(* PLC project PR_TabTrimSeq_Soft2.0 1_workflow_23a3c5_PLC, SiemensToBackhoff Siemens TIA Portal → Beckhoff TwinCAT PLCopen Converter 2.2 *)
(* stored: creationDateTime 2026-10-12T09:25:37.624382, modificationDateTime 2026-10-12T09:25:37.624382 *)

FUNCTION_BLOCK PR_TabTrimSeq_Soft2.0 1_workflow_23a3c5
VAR_INPUT
	iAbort : BOOL;
	iAutoRunning : BOOL;
	iFaultReset : BOOL;
	iPartNotWorkable : BOOL;
	iPartWorkable : BOOL;
	iRFReadDone : BOOL;
	iRFReadError : BOOL;
	iRFWriteDone : BOOL;
	iRFWriteError : BOOL;
	iReject : BOOL;
	iReset_fault : BOOL;
	iRetry : BOOL;
	iRetryCount : INT;
	iSstMode : BOOL;
	iSstPB : BOOL;
	iStartFrmFibro : BOOL;
	iStartFrmFibroSeq : BOOL;
	iTrimOver : BOOL;
	iZAxisDownOver : BOOL;
	iZAxisUpOver : BOOL;
END_VAR
VAR_OUTPUT
	qError : ARRAY[0..2] OF BOOL;
	qMessage : ARRAY[0..2] OF BOOL;
	qScrapSuction : BOOL;
	qTrimOprnOver : BOOL;
	qTrimStartCmd : BOOL;
	qZAxisUp : BOOL;
	qzAxisDown : BOOL;
END_VAR
VAR
	c20_ChkRecovery_T1 : BOOL;
	c20_ChkRecovery_T2 : BOOL;
	c20_ChkRecovery_T3 : BOOL;
	c21_WtRFIDReadOver_T1 : BOOL;
	c21_WtRFIDReadOver_T2 : BOOL;
	c22_ChkRetryCountRead_T1 : BOOL;
	c22_ChkRetryCountRead_T2 : BOOL;
	c23_WtOpDecisionRead_T1 : BOOL;
	c23_WtOpDecisionRead_T2 : BOOL;
	c24_ChkPartWorkable_T1 : BOOL;
	c24_ChkPartWorkable_T2 : BOOL;
	c61_WtRFIDWriteOver_T1 : BOOL;
	c61_WtRFIDWriteOver_T2 : BOOL;
	c62_ChkRetryCountWrite_T1 : BOOL;
	c62_ChkRetryCountWrite_T2 : BOOL;
	c63_WtOpDecisionWrite_T1 : BOOL;
	c63_WtOpDecisionWrite_T2 : BOOL;
	StateNo : INT;
	s10_WtStart : BOOL;
	s10_WtStart_T1 : BOOL;
	s1_WtResetRel : BOOL;
	s1_WtResetRel_T1 : BOOL;
	s20_ChkRecovery : BOOL;
	s20_ChkRecovery_T1 : BOOL;
	s20_ChkRecovery_T2 : BOOL;
	s20_ChkRecovery_T3 : BOOL;
	s21_WtRFIDReadOver : BOOL;
	s21_WtRFIDReadOver_T1 : BOOL;
	s21_WtRFIDReadOver_T2 : BOOL;
	s22_ChkRetryCountRead : BOOL;
	s22_ChkRetryCountRead_T1 : BOOL;
	s22_ChkRetryCountRead_T2 : BOOL;
	s23_WtOpDecisionRead : BOOL;
	s23_WtOpDecisionRead_T1 : BOOL;
	s23_WtOpDecisionRead_T2 : BOOL;
	s24_ChkPartWorkable : BOOL;
	s24_ChkPartWorkable_T1 : BOOL;
	s24_ChkPartWorkable_T2 : BOOL;
	s30_WtOperatorAck : BOOL;
	s30_WtOperatorAck_T1 : BOOL;
	s40_WtZAxisDown : BOOL;
	s40_WtZAxisDown_T1 : BOOL;
	s50_WtTrimOver : BOOL;
	s50_WtTrimOver_T1 : BOOL;
	s60_WtZAxisUp : BOOL;
	s60_WtZAxisUp_T1 : BOOL;
	s61_WtRFIDWriteOver : BOOL;
	s61_WtRFIDWriteOver_T1 : BOOL;
	s61_WtRFIDWriteOver_T2 : BOOL;
	s62_ChkRetryCountWrite : BOOL;
	s62_ChkRetryCountWrite_T1 : BOOL;
	s62_ChkRetryCountWrite_T2 : BOOL;
	s63_WtOpDecisionWrite : BOOL;
	s63_WtOpDecisionWrite_T1 : BOOL;
	s63_WtOpDecisionWrite_T2 : BOOL;
	s70_WtStartLow : BOOL;
	s70_WtStartLow_T1 : BOOL;
	sAbNormalCond : BOOL;
	sRFReadRetryCount : INT;
	sRFWriteRetryCount : INT;
	sSst : BOOL;
	sSstPulse : BOOL;
	sSstRise : R_TRIG;
	sStWtResetRel : BOOL;
	sStWtResetRel_T1 : BOOL;
	sTrimProcessActive : BOOL;
END_VAR
VAR_TEMP
	tOne : BOOL;
END_VAR
  VAR  (* added by the conversion: wires and edge detectors of the diagram *)
    _w24 : BOOL;
    _w26 : BOOL;
    _w39 : BOOL;
    _w41 : BOOL;
    _w42 : BOOL;
    _w60 : BOOL;
    _w63 : BOOL;
    _w64 : BOOL;
    _w98 : BOOL;
    _w101 : BOOL;
    _w102 : BOOL;
    _w103 : BOOL;
    _w104 : BOOL;
    _w117 : BOOL;
    _w119 : BOOL;
    _w120 : BOOL;
    _w155 : BOOL;
    _w159 : BOOL;
    _w160 : BOOL;
    _w161 : BOOL;
    _w190 : BOOL;
    _w192 : BOOL;
    _w193 : BOOL;
    _w194 : BOOL;
    _w219 : BOOL;
    _w221 : BOOL;
    _w222 : BOOL;
    _w223 : BOOL;
    _w249 : BOOL;
    _w251 : BOOL;
    _w252 : BOOL;
    _w253 : BOOL;
    _w266 : BOOL;
    _w268 : BOOL;
    _w269 : BOOL;
    _w286 : BOOL;
    _w289 : BOOL;
    _w290 : BOOL;
    _w305 : BOOL;
    _w309 : BOOL;
    _w310 : BOOL;
    _w339 : BOOL;
    _w343 : BOOL;
    _w344 : BOOL;
    _w345 : BOOL;
    _w377 : BOOL;
    _w379 : BOOL;
    _w380 : BOOL;
    _w381 : BOOL;
    _w410 : BOOL;
    _w412 : BOOL;
    _w413 : BOOL;
    _w414 : BOOL;
    _w432 : BOOL;
    _w435 : BOOL;
    _w436 : BOOL;
  END_VAR

(* LD diagram, written out as Structured Text *)
(* Network 1 *)
(* Create Single Step Pulse bit *)
(* Create Single Step bit *)
(* Transition for STATE Num:0 Reset Released *)
(* STATE Num:0 Reset Released *)
(* Transition for STATE Num:1 Wait For Reset Release *)
(* STATE Num:1 Wait For Reset Release *)
(* Transition for STATE Num:10 Wait for Start *)
(* STATE Num:10 Wait for Start *)
(* Condition1 for STATE Num:20 Check Recovery *)
(* Condition2 for STATE Num:20 Check Recovery *)
(* Condition3 for STATE Num:20 Check Recovery *)
(* Transition for STATE Num:20 Check Recovery *)
(* STATE Num:20 Check Recovery *)
(* Transition for STATE Num:30 Wait for Operator Ack *)
(* STATE Num:30 Wait for Operator Ack *)
(* Actions for STATE Num:30 Wait for Operator Ack *)
(* Condition1 for STATE Num:21 Wait for RFID Read Over *)
(* Condition2 for STATE Num:21 Wait for RFID Read Over *)
(* Transition for STATE Num:21 Wait for RFID Read Over *)
(* STATE Num:21 Wait for RFID Read Over *)
(* Condition1 for STATE Num:22 Check Retry Count Over_Read *)
(* Condition2 for STATE Num:22 Check Retry Count Over_Read *)
(* Transition for STATE Num:22 Check Retry Count Over_Read *)
(* STATE Num:22 Check Retry Count Over_Read *)
(* Condition1 for STATE Num:23 Wait For Operator decision_Read *)
(* Condition2 for STATE Num:23 Wait For Operator decision_Read *)
(* Transition for STATE Num:23 Wait For Operator decision_Read *)
(* STATE Num:23 Wait For Operator decision_Read *)
(* Condition1 for STATE Num:24 Check Part is Workable *)
(* Condition2 for STATE Num:24 Check Part is Workable *)
(* Transition for STATE Num:24 Check Part is Workable *)
(* STATE Num:24 Check Part is Workable *)
(* Transition for STATE Num:40 Wait for Z axis Down *)
(* STATE Num:40 Wait for Z axis Down *)
(* Actions for STATE Num:40 Wait for Z axis Down *)
(* Transition for STATE Num:50 Wait for Trim Over *)
(* STATE Num:50 Wait for Trim Over *)
(* Transition for STATE Num:60 Wait For Z Axis Up *)
(* STATE Num:60 Wait For Z Axis Up *)
(* Actions for STATE Num:60 Wait For Z Axis Up *)
(* Condition1 for STATE Num:61 Wait For RFID Write Over *)
(* Condition2 for STATE Num:61 Wait For RFID Write Over *)
(* Transition for STATE Num:61 Wait For RFID Write Over *)
(* STATE Num:61 Wait For RFID Write Over *)
(* Actions for STATE Num:61 Wait For RFID Write Over *)
(* Condition1 for STATE Num:62 Check Retry Count Over_Write *)
(* Condition2 for STATE Num:62 Check Retry Count Over_Write *)
(* Transition for STATE Num:62 Check Retry Count Over_Write *)
(* STATE Num:62 Check Retry Count Over_Write *)
(* Actions for STATE Num:62 Check Retry Count Over_Write *)
(* Condition1 for STATE Num:63 Wait for Operator Decision_Write *)
(* Condition2 for STATE Num:63 Wait for Operator Decision_Write *)
(* Transition for STATE Num:63 Wait for Operator Decision_Write *)
(* STATE Num:63 Wait for Operator Decision_Write *)
(* Transition for STATE Num:70 Wait For StartLow *)
(* STATE Num:70 Wait For StartLow *)
tOne := tOne OR NOT tOne;
sSstRise(CLK := iSstPB);
sSstPulse := sSstRise.Q;
sSst := iSstMode AND sSstPulse OR NOT iSstMode;
sStWtResetRel_T1 := sStWtResetRel AND iAutoRunning;
_w24 := sStWtResetRel;
_w26 := (_w24 OR NOT iAutoRunning) AND NOT sStWtResetRel_T1;
sStWtResetRel := _w26;
IF _w26 THEN StateNo := 0; END_IF;
s1_WtResetRel_T1 := s1_WtResetRel AND NOT sStWtResetRel AND sSst AND iAutoRunning;
_w39 := s1_WtResetRel;
_w41 := (_w39 OR sStWtResetRel_T1) AND NOT sStWtResetRel;
_w42 := _w41 AND NOT s1_WtResetRel_T1;
s1_WtResetRel := _w42;
IF _w42 THEN StateNo := 1; END_IF;
s10_WtStart_T1 := s10_WtStart AND NOT sStWtResetRel AND sSst AND iStartFrmFibroSeq;
IF s10_WtStart AND NOT sStWtResetRel AND sSst AND iStartFrmFibroSeq THEN sTrimProcessActive := FALSE; END_IF;
IF s10_WtStart AND NOT sStWtResetRel AND sSst AND iStartFrmFibroSeq THEN sRFReadRetryCount := 0; END_IF;
IF s10_WtStart AND NOT sStWtResetRel AND sSst AND iStartFrmFibroSeq THEN sRFWriteRetryCount := 0; END_IF;
_w60 := s10_WtStart;
_w63 := (_w60 OR s1_WtResetRel_T1 OR s70_WtStartLow_T1) AND NOT sStWtResetRel;
_w64 := _w63 AND NOT s10_WtStart_T1;
s10_WtStart := _w64;
IF _w64 THEN StateNo := 10; END_IF;
c20_ChkRecovery_T1 := sAbNormalCond;
c20_ChkRecovery_T2 := NOT sAbNormalCond AND sTrimProcessActive;
c20_ChkRecovery_T3 := NOT sAbNormalCond AND NOT sTrimProcessActive;
s20_ChkRecovery_T1 := s20_ChkRecovery AND NOT sStWtResetRel AND sSst AND c20_ChkRecovery_T1;
s20_ChkRecovery_T2 := s20_ChkRecovery AND NOT sStWtResetRel AND sSst AND NOT s20_ChkRecovery_T1 AND c20_ChkRecovery_T2;
s20_ChkRecovery_T3 := s20_ChkRecovery AND NOT sStWtResetRel AND sSst AND NOT s20_ChkRecovery_T1 AND NOT s20_ChkRecovery_T2 AND c20_ChkRecovery_T3;
_w98 := s20_ChkRecovery;
_w101 := (_w98 OR s10_WtStart_T1 OR s30_WtOperatorAck_T1) AND NOT sStWtResetRel;
_w102 := _w101 AND NOT s20_ChkRecovery_T1;
_w103 := _w102 AND NOT s20_ChkRecovery_T2;
_w104 := _w103 AND NOT s20_ChkRecovery_T3;
s20_ChkRecovery := _w104;
IF _w104 THEN StateNo := 20; END_IF;
s30_WtOperatorAck_T1 := s30_WtOperatorAck AND NOT sStWtResetRel AND sSst AND iFaultReset;
_w117 := s30_WtOperatorAck;
_w119 := (_w117 OR s20_ChkRecovery_T1) AND NOT sStWtResetRel;
_w120 := _w119 AND NOT s30_WtOperatorAck_T1;
s30_WtOperatorAck := _w120;
IF _w120 THEN StateNo := 30; END_IF;
qError[0] := s30_WtOperatorAck;
c21_WtRFIDReadOver_T1 := iRFReadError;
c21_WtRFIDReadOver_T2 := NOT iRFReadError AND iRFReadDone;
s21_WtRFIDReadOver_T1 := s21_WtRFIDReadOver AND NOT sStWtResetRel AND sSst AND c21_WtRFIDReadOver_T1;
qMessage[0] := s21_WtRFIDReadOver AND NOT sStWtResetRel AND sSst AND c21_WtRFIDReadOver_T1;
IF s21_WtRFIDReadOver AND NOT sStWtResetRel AND sSst AND c21_WtRFIDReadOver_T1 THEN sRFReadRetryCount := sRFReadRetryCount + 1; END_IF;
s21_WtRFIDReadOver_T2 := s21_WtRFIDReadOver AND NOT sStWtResetRel AND sSst AND NOT s21_WtRFIDReadOver_T1 AND c21_WtRFIDReadOver_T2;
IF s21_WtRFIDReadOver AND NOT sStWtResetRel AND sSst AND NOT s21_WtRFIDReadOver_T1 AND c21_WtRFIDReadOver_T2 THEN sRFReadRetryCount := 0; END_IF;
_w155 := s21_WtRFIDReadOver;
_w159 := (_w155 OR s20_ChkRecovery_T3 OR s22_ChkRetryCountRead_T2 OR s23_WtOpDecisionRead_T2) AND NOT sStWtResetRel;
_w160 := _w159 AND NOT s21_WtRFIDReadOver_T1;
_w161 := _w160 AND NOT s21_WtRFIDReadOver_T2;
s21_WtRFIDReadOver := _w161;
IF _w161 THEN StateNo := 21; END_IF;
c22_ChkRetryCountRead_T1 := sRFReadRetryCount > iRetryCount;
c22_ChkRetryCountRead_T2 := sRFReadRetryCount <= iRetryCount;
s22_ChkRetryCountRead_T1 := s22_ChkRetryCountRead AND NOT sStWtResetRel AND sSst AND c22_ChkRetryCountRead_T1;
qError[1] := s22_ChkRetryCountRead AND NOT sStWtResetRel AND sSst AND c22_ChkRetryCountRead_T1;
s22_ChkRetryCountRead_T2 := s22_ChkRetryCountRead AND NOT sStWtResetRel AND sSst AND NOT s22_ChkRetryCountRead_T1 AND c22_ChkRetryCountRead_T2;
_w190 := s22_ChkRetryCountRead;
_w192 := (_w190 OR s21_WtRFIDReadOver_T1) AND NOT sStWtResetRel;
_w193 := _w192 AND NOT s22_ChkRetryCountRead_T1;
_w194 := _w193 AND NOT s22_ChkRetryCountRead_T2;
s22_ChkRetryCountRead := _w194;
IF _w194 THEN StateNo := 22; END_IF;
c23_WtOpDecisionRead_T1 := iReject OR iAbort;
c23_WtOpDecisionRead_T2 := iRetry;
s23_WtOpDecisionRead_T1 := s23_WtOpDecisionRead AND NOT sStWtResetRel AND sSst AND c23_WtOpDecisionRead_T1;
s23_WtOpDecisionRead_T2 := s23_WtOpDecisionRead AND NOT sStWtResetRel AND sSst AND NOT s23_WtOpDecisionRead_T1 AND c23_WtOpDecisionRead_T2;
_w219 := s23_WtOpDecisionRead;
_w221 := (_w219 OR s22_ChkRetryCountRead_T1) AND NOT sStWtResetRel;
_w222 := _w221 AND NOT s23_WtOpDecisionRead_T1;
_w223 := _w222 AND NOT s23_WtOpDecisionRead_T2;
s23_WtOpDecisionRead := _w223;
IF _w223 THEN StateNo := 23; END_IF;
c24_ChkPartWorkable_T1 := iPartNotWorkable;
c24_ChkPartWorkable_T2 := NOT iPartNotWorkable AND iPartWorkable;
s24_ChkPartWorkable_T1 := s24_ChkPartWorkable AND NOT sStWtResetRel AND sSst AND c24_ChkPartWorkable_T1;
qMessage[2] := s24_ChkPartWorkable AND NOT sStWtResetRel AND sSst AND c24_ChkPartWorkable_T1;
s24_ChkPartWorkable_T2 := s24_ChkPartWorkable AND NOT sStWtResetRel AND sSst AND NOT s24_ChkPartWorkable_T1 AND c24_ChkPartWorkable_T2;
_w249 := s24_ChkPartWorkable;
_w251 := (_w249 OR s21_WtRFIDReadOver_T2) AND NOT sStWtResetRel;
_w252 := _w251 AND NOT s24_ChkPartWorkable_T1;
_w253 := _w252 AND NOT s24_ChkPartWorkable_T2;
s24_ChkPartWorkable := _w253;
IF _w253 THEN StateNo := 24; END_IF;
s40_WtZAxisDown_T1 := s40_WtZAxisDown AND NOT sStWtResetRel AND sSst AND iZAxisDownOver;
_w266 := s40_WtZAxisDown;
_w268 := (_w266 OR s24_ChkPartWorkable_T2) AND NOT sStWtResetRel;
_w269 := _w268 AND NOT s40_WtZAxisDown_T1;
s40_WtZAxisDown := _w269;
IF _w269 THEN StateNo := 40; END_IF;
qzAxisDown := s40_WtZAxisDown;
s50_WtTrimOver_T1 := s50_WtTrimOver AND NOT sStWtResetRel AND sSst AND iTrimOver;
_w286 := s50_WtTrimOver;
_w289 := (_w286 OR s20_ChkRecovery_T2 OR s40_WtZAxisDown_T1) AND NOT sStWtResetRel;
_w290 := _w289 AND NOT s50_WtTrimOver_T1;
s50_WtTrimOver := _w290;
qTrimStartCmd := _w290;
qScrapSuction := _w290;
IF _w290 THEN StateNo := 50; END_IF;
s60_WtZAxisUp_T1 := s60_WtZAxisUp AND NOT sStWtResetRel AND sSst AND iZAxisUpOver;
_w305 := s60_WtZAxisUp;
_w309 := (_w305 OR s24_ChkPartWorkable_T1 OR s23_WtOpDecisionRead_T1 OR s50_WtTrimOver_T1) AND NOT sStWtResetRel;
_w310 := _w309 AND NOT s60_WtZAxisUp_T1;
s60_WtZAxisUp := _w310;
IF _w310 THEN StateNo := 60; END_IF;
qZAxisUp := s60_WtZAxisUp;
c61_WtRFIDWriteOver_T1 := iRFWriteError;
c61_WtRFIDWriteOver_T2 := NOT iRFWriteError AND iRFWriteDone;
s61_WtRFIDWriteOver_T1 := s61_WtRFIDWriteOver AND NOT sStWtResetRel AND sSst AND c61_WtRFIDWriteOver_T1;
s61_WtRFIDWriteOver_T2 := s61_WtRFIDWriteOver AND NOT sStWtResetRel AND sSst AND NOT s61_WtRFIDWriteOver_T1 AND c61_WtRFIDWriteOver_T2;
_w339 := s61_WtRFIDWriteOver;
_w343 := (_w339 OR s60_WtZAxisUp_T1 OR s62_ChkRetryCountWrite_T2 OR s63_WtOpDecisionWrite_T2) AND NOT sStWtResetRel;
_w344 := _w343 AND NOT s61_WtRFIDWriteOver_T1;
_w345 := _w344 AND NOT s61_WtRFIDWriteOver_T2;
s61_WtRFIDWriteOver := _w345;
IF _w345 THEN StateNo := 61; END_IF;
qMessage[1] := s61_WtRFIDWriteOver;
c62_ChkRetryCountWrite_T1 := sRFWriteRetryCount > iRetryCount;
c62_ChkRetryCountWrite_T2 := sRFWriteRetryCount <= iRetryCount;
s62_ChkRetryCountWrite_T1 := s62_ChkRetryCountWrite AND NOT sStWtResetRel AND sSst AND c62_ChkRetryCountWrite_T1;
s62_ChkRetryCountWrite_T2 := s62_ChkRetryCountWrite AND NOT sStWtResetRel AND sSst AND NOT s62_ChkRetryCountWrite_T1 AND c62_ChkRetryCountWrite_T2;
_w377 := s62_ChkRetryCountWrite;
_w379 := (_w377 OR s61_WtRFIDWriteOver_T1) AND NOT sStWtResetRel;
_w380 := _w379 AND NOT s62_ChkRetryCountWrite_T1;
_w381 := _w380 AND NOT s62_ChkRetryCountWrite_T2;
s62_ChkRetryCountWrite := _w381;
IF _w381 THEN StateNo := 62; END_IF;
qError[2] := s62_ChkRetryCountWrite;
c63_WtOpDecisionWrite_T1 := iReject OR iAbort;
c63_WtOpDecisionWrite_T2 := iRetry;
s63_WtOpDecisionWrite_T1 := s63_WtOpDecisionWrite AND NOT sStWtResetRel AND sSst AND c63_WtOpDecisionWrite_T1;
s63_WtOpDecisionWrite_T2 := s63_WtOpDecisionWrite AND NOT sStWtResetRel AND sSst AND NOT s63_WtOpDecisionWrite_T1 AND c63_WtOpDecisionWrite_T2;
_w410 := s63_WtOpDecisionWrite;
_w412 := (_w410 OR s62_ChkRetryCountWrite_T1) AND NOT sStWtResetRel;
_w413 := _w412 AND NOT s63_WtOpDecisionWrite_T1;
_w414 := _w413 AND NOT s63_WtOpDecisionWrite_T2;
s63_WtOpDecisionWrite := _w414;
IF _w414 THEN StateNo := 63; END_IF;
s70_WtStartLow_T1 := s70_WtStartLow AND NOT sStWtResetRel AND sSst AND NOT iStartFrmFibroSeq;
IF s70_WtStartLow AND NOT sStWtResetRel AND sSst AND NOT iStartFrmFibroSeq THEN sTrimProcessActive := FALSE; END_IF;
IF s70_WtStartLow AND NOT sStWtResetRel AND sSst AND NOT iStartFrmFibroSeq THEN sRFReadRetryCount := 0; END_IF;
IF s70_WtStartLow AND NOT sStWtResetRel AND sSst AND NOT iStartFrmFibroSeq THEN sRFWriteRetryCount := 0; END_IF;
_w432 := s70_WtStartLow;
_w435 := (_w432 OR s61_WtRFIDWriteOver_T2 OR s63_WtOpDecisionWrite_T1) AND NOT sStWtResetRel;
_w436 := _w435 AND NOT s70_WtStartLow_T1;
qTrimOprnOver := _w436;
s70_WtStartLow := _w436;
IF _w436 THEN StateNo := 70; END_IF;
END_FUNCTION_BLOCK
